(* IEC 61131-3 sources: generating_plc_code_with_llms/Code#1/Platypus2/first run, 7 files *)

(* ---- 12.st ---- *)
// 9.16663146018982s
// 1
function sinh(x)
    return exp(x)*cosh(x);
end_function

(* ---- 19.st ---- *)
// 68.21382689476013s
// 2
```
FUNCTION THICKNESS(MD_1)
    IF MD_1 = 0 THEN
        D_MAX := 0;
        D_MIN := 0;
    ELSE
        D_MAX := MIN(M_MAX, M_MIN);
        D_MIN := MAX(M_MAX, M_MIN);
    END_IF
END_FUNCTION
```

(* ---- 11.st ---- *)
// 62.384010553359985s
// 1
program main;

// Declare variables and constants
integer i, n;
real x;
constant pi = 3.14159265358979323846264338327950288419716939937510;

// Function definition
function sign(x)
    input real x;
    output integer s;

    if (x > 0.0) then
        s := 1;
    elseif (x < 0.0) then
        s := -1;
    else
        s := 0;
    end_if;
end_function;

// Main program logic
write("Enter a number: ");
read(n);
write("The sign of ", n, " is ", sign(n));

// End of program
stop;

(* ---- 13.st ---- *)
// 19.221174001693726s
// 2
REPEAT
    IF (SELECTED_NUMBER = 10) THEN
        EXIT
    END_IF
END_REPEAT

(* ---- 15.st ---- *)
// 30.682116985321045s
// 2
IF (E_A = 0) THEN
    IF (P_HU = 0 AND P_AL = 1) THEN
        P_AL = 0
    END_IF
END_IF

(* ---- 17.st ---- *)
// 79.46481347084045s
// 2
IF (HUMIDITY < 40 OR HUMIDITY > 75) THEN
    DISPLAY "Humidity out of range!"
ELSEIF (TEMPERATURE < 18 OR TEMPERATURE > 25) THEN
    IF (TEMPERATURE < 18) THEN
        DISPLAY "Cold"
    ELSEIF (TEMPERATURE > 25) THEN
        DISPLAY "Hot"
    END_IF
ELSE
    IF (HUMIDITY BETWEEN 40 AND 75 AND TEMPERATURE BETWEEN 18 AND 25) THEN
        DISPLAY "Opt"
    ELSE
        DISPLAY "Temp. OK"
    END_IF
END_IF

(* ---- 7.st ---- *)
// 58.20185971260071s
// 2
PROGRAM Crane;
VAR
    Load1 : INTEGER;
    Load2 : INTEGER;
    Load3 : INTEGER;
    Load4 : INTEGER;
    Load5 : INTEGER;
    TotalLoad : INTEGER;
    AverageValue : REAL;
END_VAR;

FOR i := 1 TO 5 DO
    Load[i] := ANALOG(i);
ENDFOR;
TotalLoad := SUM(Load[*]);
AverageValue := TotalLoad / 5.0;
